FUNCTION_BLOCK ALR_TO_ATM_IN_S (* Convert LREAL (via ALR adapter) in S to TIME (via ATM adapter), Gegenrichtung zu ATM_IN_S_TO_ALR *)
  (* Standard: 61499-2; Function: OUT = T#1s * IN (F_MULTIME); Description: Copyright (c) 2026 HR Agrartechnik GmbH This program and the accompanying materials are made available under the terms of the Eclipse Public License 2.0 which is available at https://www.eclipse.org/legal/epl-2.0/ SPDX-License-Identifier: EPL-2.0 *)
  (* Version 1.0, 2026-11-13, Franz Höpfinger, HR Agrartechnik GmbH, Initial Version - Luecke in der Adapter-Familie geschlossen *)
  PACKAGE adapter::conversion::unidirectional;
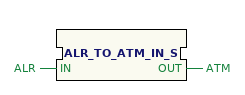
  SOCKETS
    IN : adapter::types::unidirectional::ALR; (* Zeitwert in S als LREAL *)
  END_SOCKETS
  PLUGS
    OUT : adapter::types::unidirectional::ATM; (* TIME-Wert = IN * 1 S *)
  END_PLUGS
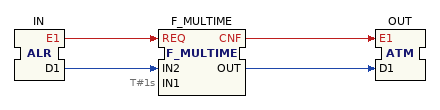
  FBS
    F_MULTIME : iec61131::arithmetic::F_MULTIME(IN1 := T#1s);
  END_FBS
  EVENT_CONNECTIONS
    IN.E1 TO F_MULTIME.REQ;
    F_MULTIME.CNF TO OUT.E1;
  END_CONNECTIONS
  DATA_CONNECTIONS
    IN.D1 TO F_MULTIME.IN2;
    F_MULTIME.OUT TO OUT.D1;
  END_CONNECTIONS
END_FUNCTION_BLOCK
